SYSTEM System
  DEVICE DEV : Soft_dPAC
    RESOURCE RES0 : EMB_RES_ECO
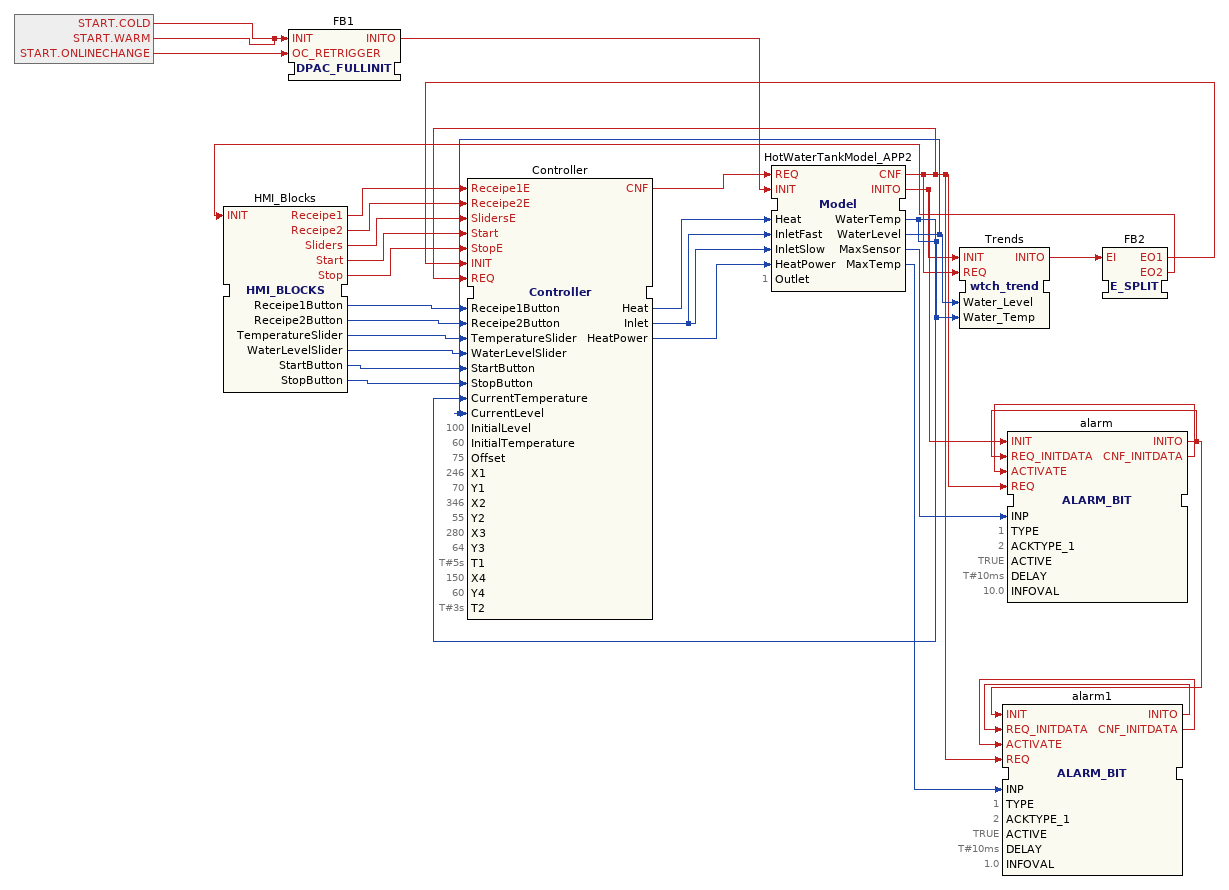
      FBS
        HotWaterTankModel_APP2 : Model(Outlet := 1);
        HMI_Blocks : HMI_BLOCKS;
        Controller : Controller(InitialLevel := 100, InitialTemperature := 60, Offset := 75, X1 := 246, Y1 := 70, X2 := 346, Y2 := 55, X3 := 280, Y3 := 64, T1 := T#5s, X4 := 150, Y4 := 60, T2 := T#3s);
        FB2 : E_SPLIT;
        Trends : wtch_trend;
        FB1 : DPAC_FULLINIT;
        alarm : ALARM_BIT(TYPE := 1, ACKTYPE_1 := 2, ACTIVE := TRUE, DELAY := T#10ms, INFOVAL := 10.0);
        alarm1 : ALARM_BIT(TYPE := 1, ACKTYPE_1 := 2, ACTIVE := TRUE, DELAY := T#10ms, INFOVAL := 1.0);
      END_FBS
      EVENT_CONNECTIONS
        HMI_Blocks.Receipe1 TO Controller.Receipe1E;
        HMI_Blocks.Receipe2 TO Controller.Receipe2E;
        HMI_Blocks.Sliders TO Controller.SlidersE;
        HMI_Blocks.Start TO Controller.Start;
        HMI_Blocks.Stop TO Controller.StopE;
        Trends.INITO TO FB2.EI;
        FB2.EO1 TO Controller.INIT;
        FB2.EO2 TO HMI_Blocks.INIT;
        Controller.CNF TO HotWaterTankModel_APP2.REQ;
        HotWaterTankModel_APP2.CNF TO Controller.REQ;
        HotWaterTankModel_APP2.INITO TO Trends.INIT;
        HotWaterTankModel_APP2.CNF TO Trends.REQ;
        START.COLD TO FB1.INIT;
        START.WARM TO FB1.INIT;
        START.ONLINECHANGE TO FB1.OC_RETRIGGER;
        FB1.INITO TO HotWaterTankModel_APP2.INIT;
        HotWaterTankModel_APP2.INITO TO alarm.INIT;
        alarm.INITO TO alarm.REQ_INITDATA;
        alarm.CNF_INITDATA TO alarm.ACTIVATE;
        HotWaterTankModel_APP2.CNF TO alarm.REQ;
        alarm.INITO TO alarm1.INIT;
        alarm1.INITO TO alarm1.REQ_INITDATA;
        alarm1.CNF_INITDATA TO alarm1.ACTIVATE;
        HotWaterTankModel_APP2.CNF TO alarm1.REQ;
      END_CONNECTIONS
      DATA_CONNECTIONS
        HMI_Blocks.Receipe1Button TO Controller.Receipe1Button;
        HMI_Blocks.Receipe2Button TO Controller.Receipe2Button;
        HMI_Blocks.TemperatureSlider TO Controller.TemperatureSlider;
        HMI_Blocks.WaterLevelSlider TO Controller.WaterLevelSlider;
        HMI_Blocks.StartButton TO Controller.StartButton;
        HMI_Blocks.StopButton TO Controller.StopButton;
        Controller.Heat TO HotWaterTankModel_APP2.Heat;
        Controller.Inlet TO HotWaterTankModel_APP2.InletFast;
        Controller.Inlet TO HotWaterTankModel_APP2.InletSlow;
        HotWaterTankModel_APP2.WaterTemp TO Controller.CurrentTemperature;
        HotWaterTankModel_APP2.WaterLevel TO Controller.CurrentLevel;
        Controller.HeatPower TO HotWaterTankModel_APP2.HeatPower;
        HotWaterTankModel_APP2.WaterLevel TO Trends.Water_Level;
        HotWaterTankModel_APP2.WaterTemp TO Trends.Water_Temp;
        HotWaterTankModel_APP2.MaxSensor TO alarm.INP;
        HotWaterTankModel_APP2.MaxTemp TO alarm1.INP;
      END_CONNECTIONS
    END_RESOURCE
  END_DEVICE
END_SYSTEM
